(* IEC 61131-3 sources: 2026_Projet_YGO_ExcavatriceDragage/ARCHIVES/Code/CFC_STAGING_RECOVERED/CODE/TRANSLATION, 5 files *)

(* ---- FB_TranslationArbiter.st ---- *)
(* ═══════════════════════════════════════════════════════════════
   ↔️ FB_TranslationArbiter — Arbitrage des consignes M3
   ───────────────────────────────────────────────────────────────
   📄 Migration M4 : extrait sans changement la logique de page de
      PRG_TRANSLATION_CFC.st afin que le CFC natif ne porte aucun IF/CASE.
   🔒 Ce FB ne commande aucun actionneur : il produit uniquement la demande
      arbitrée consommée par FB_Translation.
   ═══════════════════════════════════════════════════════════════ *)

FUNCTION_BLOCK PUBLIC FB_TranslationArbiter
VAR_INPUT
    Mode                         : E_Mode;
    AutoStart                    : BOOL;
    AutoTarget                   : INT;
    DeadmanArmed                 : BOOL;
    AxisCmd                      : ST_Joystick_AxisCmd;
    MaintenancePositioning       : BOOL;
    MaintenanceTarget            : INT;
    BtnFwd                       : BOOL;
    BtnRev                       : BOOL;
    TglJoystickMaster            : BOOL;
    SetFreqHz                    : REAL;
    BypassGlobal                 : BOOL;
    InvertDirection              : BOOL;
    MaintenanceM3TargetEnable    : BOOL;
    PosTremie                    : BOOL;
    PosP2                        : BOOL;
    PosP1                        : BOOL;
    PosMaintenance               : BOOL;
    AutoSpeedCapPct              : REAL;
    TranslationMaxFreqHz         : REAL;
END_VAR
VAR_OUTPUT
    StartStop                    : BOOL;
    Direction                    : INT;
    SpeedRefPct                  : REAL;
    PositionSensorTarget         : BOOL;
    PositioningActive            : BOOL;
    SelectedTarget               : INT;
END_VAR
VAR
    FreqPct                      : REAL;
END_VAR

(* ── Arbitrage sources Semi-auto / Maintenance / conduite manuelle ── *)
IF Mode = E_Mode.SEMI_AUTO THEN
    PositioningActive := TRUE;
    SelectedTarget := AutoTarget;
    StartStop := AutoStart AND DeadmanArmed AND AxisCmd.StartStop;
    SpeedRefPct := ABS(AxisCmd.SpeedRef);
    IF SpeedRefPct > AutoSpeedCapPct THEN
        SpeedRefPct := AutoSpeedCapPct;
    END_IF;

    IF SelectedTarget = 1 THEN
        Direction := 1;
    ELSE
        Direction := -1;
    END_IF;
ELSIF (Mode = E_Mode.MAINT_N1) OR (Mode = E_Mode.MAINT_N2) THEN
    PositioningActive := MaintenancePositioning;
    IF PositioningActive THEN
        SelectedTarget := MaintenanceTarget;
    ELSE
        SelectedTarget := 0;
    END_IF;

    IF (NOT TglJoystickMaster) AND BtnFwd THEN
        Direction := 1;
    ELSIF (NOT TglJoystickMaster) AND BtnRev THEN
        Direction := -1;
    ELSIF TglJoystickMaster THEN
        Direction := AxisCmd.Direction;
    ELSE
        Direction := 0;
    END_IF;

    StartStop := (Direction <> 0)
                 AND (DeadmanArmed OR BypassGlobal)
                 AND ((NOT TglJoystickMaster) OR AxisCmd.StartStop);

    IF SetFreqHz > 0.0 THEN
        FreqPct := (SetFreqHz / TranslationMaxFreqHz) * 100.0;
    ELSE
        FreqPct := 30.0;
    END_IF;

    IF TglJoystickMaster THEN
        SpeedRefPct := (ABS(AxisCmd.SpeedRef) / 100.0) * FreqPct;
    ELSE
        SpeedRefPct := FreqPct;
    END_IF;
ELSE
    PositioningActive := FALSE;
    SelectedTarget := MaintenanceTarget;
    StartStop := AxisCmd.StartStop;
    Direction := AxisCmd.Direction;
    SpeedRefPct := AxisCmd.SpeedRef;
END_IF;

(* ── Gardes conservation : inversion, borne vitesse, MAINT_N2 et cible ── *)
IF InvertDirection THEN
    Direction := Direction * (-1);
END_IF;

SpeedRefPct := ABS(SpeedRefPct);
IF SpeedRefPct > 100.0 THEN
    SpeedRefPct := 100.0;
END_IF;

IF (SelectedTarget = 4) AND (NOT MaintenanceM3TargetEnable) THEN
    SelectedTarget := 0;
END_IF;

CASE SelectedTarget OF
    1: PositionSensorTarget := PosTremie;
    2: PositionSensorTarget := PosP2;
    3: PositionSensorTarget := PosP1;
    4: PositionSensorTarget := PosMaintenance;
ELSE
    PositionSensorTarget := FALSE;
END_CASE;

(* ---- FB_TranslationCfcExpressions.st ---- *)
(* ═══════════════════════════════════════════════════════════════
   ↔️ FB_TranslationCfcExpressions — Expressions extraites du CFC
   ───────────────────────────────────────────────────────────────
   🎯 Rôle : porter les trois expressions booléennes du câblage
      historique dans un FB ST, afin que la page CFC XML ne comporte
      que des blocs et des fils.

   🔒 Conservation : chaque sortie est l'expression legacy à l'identique.
   Aucun accès sortie physique, aucune décision de sécurité nouvelle.
   ═══════════════════════════════════════════════════════════════ *)
FUNCTION_BLOCK FB_TranslationCfcExpressions
VAR_INPUT
    BrakeThermalFeedback       : BOOL;
    BypassContactorFeedback    : BOOL;
    BypassGlobal               : BOOL;
    BypassLimitSwitch          : BOOL;
END_VAR
VAR_OUTPUT
    BrakeThermalOk                 : BOOL;
    BypassContactorFeedbackEffective : BOOL;
    BypassLimitSwitchEffective       : BOOL;
END_VAR

BrakeThermalOk := NOT BrakeThermalFeedback;
BypassContactorFeedbackEffective := BypassContactorFeedback OR BypassGlobal;
BypassLimitSwitchEffective := BypassGlobal OR BypassLimitSwitch;

(* ---- FB_TranslationFeedbackMemory.st ---- *)
(* ═══════════════════════════════════════════════════════════════
   ↔️ FB_TranslationFeedbackMemory — Mémoire N-1 desserrage frein M3
   ───────────────────────────────────────────────────────────────
   📄 Migration M4 : rend explicite la lecture historique du propre
      BrakeReleaseRequest de instTranslationM3 avant son appel du scan.
   🔒 Cette mémoire ne prouve pas la position mécanique du frein. Le retour
      physique reste BrakeFeedback; la dette BrakeCmd A-07 reste inchangée.
   ═══════════════════════════════════════════════════════════════ *)

FUNCTION_BLOCK PUBLIC FB_TranslationFeedbackMemory
VAR_INPUT
    BrakeReleaseRequest : BOOL;
END_VAR
VAR_OUTPUT
    PreviousBrakeReleaseRequest : BOOL;
END_VAR
VAR
    StoredBrakeReleaseRequest : BOOL := FALSE;
END_VAR

PreviousBrakeReleaseRequest := StoredBrakeReleaseRequest;
StoredBrakeReleaseRequest := BrakeReleaseRequest;

(* ---- FB_TranslationRequestPublisher.st ---- *)
(* ═══════════════════════════════════════════════════════════════
   ↔️ FB_TranslationRequestPublisher — Contrat M3 vers Outputs
   ───────────────────────────────────────────────────────────────
   📄 Migration M4 : encapsule l'assemblage de
      ST_TranslationFinalInterlockRequest hors de la page CFC native.
   🔒 Ne produit qu'une demande brute; PRG_06_Outputs_LD reste l'unique
      propriétaire des commandes physiques AC600 et du frein.
   ═══════════════════════════════════════════════════════════════ *)

FUNCTION_BLOCK PUBLIC FB_TranslationRequestPublisher
VAR_INPUT
    Enable                      : BOOL;
    Reset                       : BOOL;
    PowerContactorEngaged       : BOOL;
    SafeStop                    : BOOL;
    BrakeReleaseRequest         : BOOL;
    BrakeCommandOpenConfirmed   : BOOL;
    RequestedDriveControlWord   : WORD;
    RequestedDriveFreqHz        : REAL;
END_VAR
VAR_OUTPUT
    Request                     : ST_TranslationFinalInterlockRequest;
END_VAR

Request.Enable := Enable;
Request.Reset := Reset;
Request.PowerContactorEngaged := PowerContactorEngaged;
Request.SafeStop := SafeStop;
Request.BrakeReleaseRequest := BrakeReleaseRequest;
Request.BrakeCommandOpenConfirmed := BrakeCommandOpenConfirmed;
Request.RequestedDriveControlWord := RequestedDriveControlWord;
Request.RequestedDriveFreqHz := RequestedDriveFreqHz;

(* ---- FB_TranslationRuntimeGate.st ---- *)
(* ═══════════════════════════════════════════════════════════════
   ↔️ FB_TranslationRuntimeGate — Préconditions d'appel FB_Translation
   ───────────────────────────────────────────────────────────────
   📄 Migration M4 : extrait les expressions booléennes/SEL de la page
      historique pour conserver un CFC XML sans calcul inline.
   🔒 Le retour de desserrage est lu à N-1 via FB_TranslationFeedbackMemory,
      identique à l'auto-référence historique instTranslationM3.BrakeReleaseRequest.
   ═══════════════════════════════════════════════════════════════ *)

FUNCTION_BLOCK PUBLIC FB_TranslationRuntimeGate
VAR_INPUT
    MachineEnable                 : BOOL;
    Mode                          : E_Mode;
    BypassContactorFeedback       : BOOL;
    BrakeFeedback                 : BOOL;
    PreviousBrakeReleaseRequest   : BOOL;
END_VAR
VAR_OUTPUT
    Enable                        : BOOL;
    BrakeFeedbackForTranslation   : BOOL;
END_VAR

Enable := MachineEnable AND (Mode <> E_Mode.DISABLE);

IF BypassContactorFeedback THEN
    BrakeFeedbackForTranslation := PreviousBrakeReleaseRequest;
ELSE
    BrakeFeedbackForTranslation := BrakeFeedback;
END_IF;
